TYPE ST_PERIPHERY_REF_1 : FB_PERIPHERY_REF;
END_TYPE

(* stored: Version 1.1.0.1, ProductVersion 3.1.4024.15
   DUT ST_PERIPHERY_REF_1: Id {2ccfff72-37d8-4de5-b12d-498bed54a070} *)
